TYPE TcoKukaKss_Outputs_v_9_3_x :
STRUCT
	Outputs AT %Q* : ARRAY[0..63] OF BYTE;
END_STRUCT
END_TYPE

(* stored: Version 1.1.0.1, ProductVersion 3.1.4024.12
   DUT TcoKukaKss_Outputs_v_9_3_x: Id {af8bca6f-ef4c-4fd6-bf22-ccbbadf99a85} *)
